Fanuc KAREL source: KD00003.KL

PROGRAM KD00003
%NOLOCKGROUP
%CMOSVARS
VAR
  I: INTEGER
  J: INTEGER
  B: BOOLEAN
  R: REAL
  S: STRING[80]
BEGIN
  I = 1
END KD00003
